(* IEC 61131-3 sources: codesys_asrs/Project_ASRS_CodeSYS (part 2) *)

(* ---- 16_FB_G3_Cycle_BODY_ONLY.st ---- *)
T_Nettoyage15(IN := NettoyageTimerEnable AND NOT GVL_SIG.ZONE_CONFIRMEE, PT := T#15m);
T_Prolong5(IN := ProlongTimerEnable AND NOT GVL_SIG.ZONE_CONFIRMEE, PT := T#5m);

// â”€â”€ Surveillance AU pendant cycle (prioritÃ© absolue) â”€â”€â”€â”€â”€â”€â”€â”€â”€â”€
IF GVL_SIG.OP_AU AND Step > 0 AND Step < 200 THEN
    GVL_SIG.G3_DEFAUT      := TRUE;
    GVL_SIG.G3_CODE_DEFAUT := 14;
    GVL_SEQ.DEFAUT_ACTIF   := TRUE;
    GVL_SEQ.CODE_DEFAUT    := 14;
    GVL_SIG.G4_REQ         := FALSE;
    GVL_SIG.G5_REQ         := FALSE;
    GVL_SIG.G6_REQ         := FALSE;
    GVL_SIG.G7_REQ         := FALSE;
    GVL_SIG.G8_REQ         := FALSE;
    GVL_SIG.G9_REQ_ARRET     := FALSE;
    GVL_SIG.G10_REQ_ENTRER   := FALSE;
    GVL_SIG.G10_REQ_SORTIR   := FALSE;
    GVL_SIG.VYT_CYCLE_EN_COURS := FALSE;
    Step := 0;
    RETURN;
END_IF;

CASE Step OF

// â•â•â•â•â•â•â•â•â•â•â•â•â•â•â•â•â•â•â•â•â•â•â•â•â•â•â•â•â•â•â•â•â•â•â•â•â•â•â•â•â•â•â•â•â•â•â•â•â•â•â•â•â•â•â•â•â•â•â•â•
// PHASE 0 â€” IDLE
// â•â•â•â•â•â•â•â•â•â•â•â•â•â•â•â•â•â•â•â•â•â•â•â•â•â•â•â•â•â•â•â•â•â•â•â•â•â•â•â•â•â•â•â•â•â•â•â•â•â•â•â•â•â•â•â•â•â•â•â•
0:
    GVL_SIG.G3_FIN_CM          := FALSE;
    GVL_SIG.G3_DEFAUT          := FALSE;
    GVL_SIG.G3_CODE_DEFAUT     := 0;
    GVL_SIG.VYT_CYCLE_EN_COURS := FALSE;
    GVL_SIG.G9_ARRETEE_OK      := FALSE;
    GVL_SIG.G9_DEBRIDE_OK      := FALSE;
    GVL_SIG.G9_BRIDE_OK        := FALSE;
    GVL_SIG.G9_AUTORISE_OK     := FALSE;
    GVL_SIG.G10_EN_PRESSE      := FALSE;
    GVL_SIG.G10_A_ZPM          := FALSE;
    NettoyageTimerEnable       := FALSE;
    ProlongTimerEnable         := FALSE;
    GVL_SIG.NETTOYAGE_EN_COURS := FALSE;
    GVL_SIG.NETTOYAGE_TIMEOUT  := FALSE;
    GVL_SIG.NETTOYAGE_PROLONGATION_UTILISEE := FALSE;
    GVL_SIG.NETTOYAGE_DEPASSEMENT_MAX := FALSE;
    GVL_SIG.VYT_NETTOYAGE_TIMEOUT := FALSE;
    GVL_IO.VOYANT_NETTOYAGE_TIMEOUT := FALSE;
    GVL_IO.VOYANT_NETTOYAGE_MAX := FALSE;
    GVL_IO.BUZZER_ATTENTE_ZONE_LIBRE := FALSE;
    IF GVL_SIG.G3_REQ THEN
        DepotFound := FALSE;
        PriseFound := FALSE;
        IF GVL_MOULES.MOULE_EN_PRESSE = 0 THEN
            GVL_SIG.G3_CODE_DEFAUT := 16;
            Step := 200;
        ELSIF GVL_MOULES.MOULE_DEMANDE = 0 THEN
            GVL_SIG.G3_CODE_DEFAUT := 13;
            Step := 200;
        ELSIF GVL_MOULES.MOULE_DEMANDE = GVL_MOULES.MOULE_EN_PRESSE THEN
            GVL_SIG.G3_CODE_DEFAUT := 17;
            Step := 200;
        ELSE
            Step := 1;
        END_IF;
    END_IF;

1: // Recherche slot dÃ©pÃ´t
    DepotFound := FALSE;
    FOR i := 1 TO 5 BY 1 DO
        IF NOT DepotFound THEN
            FOR j := 1 TO 2 BY 1 DO
                IF NOT DepotFound
                   AND NOT GVL_MOULES.CH[i, j].OCCUPE
                   AND NOT GVL_MOULES.CH[i, j].RESERVE THEN
                    GVL_MOULES.CIBLE_DEPOT_CH := INT_TO_USINT(i);
                    GVL_MOULES.CIBLE_DEPOT_NV := INT_TO_USINT(j);
                    GVL_MOULES.CH[i, j].RESERVE := TRUE;
                    DepotFound := TRUE;
                END_IF;
            END_FOR;
        END_IF;
    END_FOR;
    IF DepotFound THEN
        Step := 2;
    ELSE
        GVL_MOULES.ALM_STOCK_PLEIN := TRUE;
        GVL_SIG.ALM_STOCK_PLEIN   := TRUE;
        GVL_SIG.G3_CODE_DEFAUT    := 12;
        Step := 200;
    END_IF;

2: // Recherche slot prise
    PriseFound := FALSE;
    FOR i := 1 TO 5 BY 1 DO
        IF NOT PriseFound THEN
            FOR j := 1 TO 2 BY 1 DO
                IF NOT PriseFound
                   AND GVL_MOULES.CH[i, j].OCCUPE
                   AND GVL_MOULES.CH[i, j].ID = GVL_MOULES.MOULE_DEMANDE THEN
                    GVL_MOULES.CIBLE_PRISE_CH := INT_TO_USINT(i);
                    GVL_MOULES.CIBLE_PRISE_NV := INT_TO_USINT(j);
                    PriseFound := TRUE;
                END_IF;
            END_FOR;
        END_IF;
    END_FOR;
    IF PriseFound THEN
        GVL_SIG.VYT_CYCLE_EN_COURS := TRUE;
        Step := 3;
    ELSE
        GVL_MOULES.CH[GVL_MOULES.CIBLE_DEPOT_CH, GVL_MOULES.CIBLE_DEPOT_NV].RESERVE := FALSE;
        GVL_SIG.G3_CODE_DEFAUT := 13;
        Step := 200;
    END_IF;

3:
    GVL_SEQ.CYCLE_INTERROMPU := TRUE;
    GVL_SEQ.CYCLE_EN_COURS   := TRUE;

// â•â•â•â•â•â•â•â•â•â•â•â•â•â•â•â•â•â•â•â•â•â•â•â•â•â•â•â•â•â•â•â•â•â•â•â•â•â•â•â•â•â•â•â•â•â•â•â•â•â•â•â•â•â•â•â•â•â•â•â•
// PHASE 1 â€” ArrÃªt presse + dÃ©bridage
// â•â•â•â•â•â•â•â•â•â•â•â•â•â•â•â•â•â•â•â•â•â•â•â•â•â•â•â•â•â•â•â•â•â•â•â•â•â•â•â•â•â•â•â•â•â•â•â•â•â•â•â•â•â•â•â•â•â•â•â•
10:
    GVL_SIG.G9_REQ_ARRET   := TRUE;
    GVL_SIG.G10_REQ_ENTRER := TRUE;
    Step := 11;

11:
    IF GVL_SIG.G9_ARRETEE_OK THEN
        GVL_SIG.G9_REQ_DEBRIDAGE := TRUE;
        Step := 12;
    ELSIF GVL_SIG.G9_DEFAUT THEN
        Step := 200;
    END_IF;

12:
    IF GVL_SIG.G9_DEBRIDE_OK THEN
        Step := 13;
    ELSIF GVL_SIG.G9_DEFAUT THEN
        Step := 200;
    END_IF;

// â•â•â•â•â•â•â•â•â•â•â•â•â•â•â•â•â•â•â•â•â•â•â•â•â•â•â•â•â•â•â•â•â•â•â•â•â•â•â•â•â•â•â•â•â•â•â•â•â•â•â•â•â•â•â•â•â•â•â•â•
// DIVERGENCE ET#1 â€” Retrait introducteur â€– Chariot â†’ P0
// â•â•â•â•â•â•â•â•â•â•â•â•â•â•â•â•â•â•â•â•â•â•â•â•â•â•â•â•â•â•â•â•â•â•â•â•â•â•â•â•â•â•â•â•â•â•â•â•â•â•â•â•â•â•â•â•â•â•â•â•
13:
    BrA_Done := FALSE;
    BrB_Done := FALSE;
    SubA     := 0;
    SubB     := 0;
    Step     := 14;

14:
    IF NOT BrA_Done THEN
        CASE SubA OF
        0:  GVL_SIG.G10_REQ_SORTIR := TRUE;
            SubA := 1;
        1:  IF GVL_SIG.G10_A_ZPM THEN
                BrA_Done := TRUE;
            ELSIF GVL_SIG.G10_DEFAUT THEN
                GVL_SIG.G3_CODE_DEFAUT := 5;
                Step := 200;
            END_IF;
        END_CASE;
    END_IF;

    IF NOT BrB_Done THEN
        CASE SubB OF
        0:  GVL_SIG.G4_REQ   := TRUE;
            GVL_SIG.G4_CIBLE := 0;
            SubB := 1;
        1:  IF GVL_SIG.G4_DONE THEN
                GVL_SIG.G4_DONE := FALSE;
                BrB_Done := TRUE;
            ELSIF GVL_SIG.G4_ERR THEN
                GVL_SIG.G4_ERR := FALSE;
                GVL_SIG.G3_CODE_DEFAUT := 7;
                Step := 200;
            END_IF;
        END_CASE;
    END_IF;

    IF BrA_Done AND BrB_Done THEN
        GVL_SIG.G10_REQ_ENTRER := FALSE;
        GVL_SIG.G10_REQ_SORTIR := FALSE;
        Step := 15;
    END_IF;

// â•â•â•â•â•â•â•â•â•â•â•â•â•â•â•â•â•â•â•â•â•â•â•â•â•â•â•â•â•â•â•â•â•â•â•â•â•â•â•â•â•â•â•â•â•â•â•â•â•â•â•â•â•â•â•â•â•â•â•â•
// PHASE 2 â€” Transfert moule : introducteur â†’ chariot
// â•â•â•â•â•â•â•â•â•â•â•â•â•â•â•â•â•â•â•â•â•â•â•â•â•â•â•â•â•â•â•â•â•â•â•â•â•â•â•â•â•â•â•â•â•â•â•â•â•â•â•â•â•â•â•â•â•â•â•â•
15:
    IF NOT GVL_IO.MOULE_SUR_INTRO THEN
        GVL_SIG.G3_CODE_DEFAUT := 13;
        Step := 200;
    ELSE
        Step := 16;
    END_IF;

16:
    GVL_SIG.G6_REQ   := TRUE;
    GVL_SIG.G6_CIBLE := 0;  // NORD
    Step := 17;

17:
    IF GVL_SIG.G6_DONE THEN
        GVL_SIG.G6_DONE := FALSE;
        Step := 18;
    ELSIF GVL_SIG.G6_ERR THEN
        GVL_SIG.G6_ERR         := FALSE;
        GVL_SIG.G3_CODE_DEFAUT := 11;
        Step := 200;
    END_IF;

18:
    GVL_SIG.G5_REQ   := TRUE;
    GVL_SIG.G5_CIBLE := 0;  // Z_ZPM
    Step := 19;

19:
    IF GVL_SIG.G5_DONE THEN
        GVL_SIG.G5_DONE := FALSE;
        Step := 20;
    ELSIF GVL_SIG.G5_ERR THEN
        GVL_SIG.G5_ERR         := FALSE;
        GVL_SIG.G3_CODE_DEFAUT := 6;
        Step := 200;
    END_IF;

20:
    GVL_SIG.G7_REQ := TRUE;
    GVL_SIG.G7_CMD := 0;  // ETENDRE
    Step := 21;

21:
    IF GVL_SIG.G7_DONE THEN
        GVL_SIG.G7_DONE := FALSE;
        Step := 22;
    ELSIF GVL_SIG.G7_ERR THEN
        GVL_SIG.G7_ERR         := FALSE;
        GVL_SIG.G3_CODE_DEFAUT := 11;
        Step := 200;
    END_IF;

22:
    GVL_SIG.G5_REQ   := TRUE;
    GVL_SIG.G5_CIBLE := 3;  // Z_TRANSPORT
    Step := 23;

23:
    IF GVL_SIG.G5_DONE THEN
        GVL_SIG.G5_DONE := FALSE;
        IF NOT GVL_IO.CAPTEUR_CHARGE_CHARIOT THEN
            GVL_SIG.G3_CODE_DEFAUT := 10;
            Step := 200;
        ELSE
            Step := 24;
        END_IF;
    ELSIF GVL_SIG.G5_ERR THEN
        GVL_SIG.G5_ERR         := FALSE;
        GVL_SIG.G3_CODE_DEFAUT := 6;
        Step := 200;
    END_IF;

24:
    GVL_SIG.G7_REQ := TRUE;
    GVL_SIG.G7_CMD := 1;  // RETRACTER
    Step := 25;

25:
    IF GVL_SIG.G7_DONE THEN
        GVL_SIG.G7_DONE := FALSE;
        Step := 26;
    ELSIF GVL_SIG.G7_ERR THEN
        GVL_SIG.G7_ERR         := FALSE;
        GVL_SIG.G3_CODE_DEFAUT := 11;
        Step := 201;
    END_IF;

// â•â•â•â•â•â•â•â•â•â•â•â•â•â•â•â•â•â•â•â•â•â•â•â•â•â•â•â•â•â•â•â•â•â•â•â•â•â•â•â•â•â•â•â•â•â•â•â•â•â•â•â•â•â•â•â•â•â•â•â•
// DIVERGENCE ET#2 â€” Stockage+RFID+Prise â€– Nettoyage
// â•â•â•â•â•â•â•â•â•â•â•â•â•â•â•â•â•â•â•â•â•â•â•â•â•â•â•â•â•â•â•â•â•â•â•â•â•â•â•â•â•â•â•â•â•â•â•â•â•â•â•â•â•â•â•â•â•â•â•â•
26:
    BrA_Done := FALSE;
    BrB_Done := FALSE;
    SubA     := 0;
    SubB     := 0;
    NettoyageTimerEnable := FALSE;
    ProlongTimerEnable := FALSE;
    GVL_SIG.NETTOYAGE_EN_COURS := FALSE;
    GVL_SIG.NETTOYAGE_TIMEOUT := FALSE;
    GVL_SIG.NETTOYAGE_PROLONGATION_UTILISEE := FALSE;
    GVL_SIG.NETTOYAGE_DEPASSEMENT_MAX := FALSE;
    GVL_SIG.VYT_NETTOYAGE_TIMEOUT := FALSE;
    GVL_IO.VOYANT_NETTOYAGE_TIMEOUT := FALSE;
    GVL_IO.VOYANT_NETTOYAGE_MAX := FALSE;
    GVL_IO.BUZZER_ATTENTE_ZONE_LIBRE := FALSE;
    Step     := 27;

27: // ET#2
    IF NOT BrA_Done THEN
        CASE SubA OF
        0:  GVL_SIG.G4_REQ   := TRUE;
            GVL_SIG.G4_CIBLE := GVL_MOULES.CIBLE_DEPOT_CH;
            SubA := 1;
        1:  IF GVL_SIG.G4_DONE THEN
                GVL_SIG.G4_DONE := FALSE; SubA := 2;
            ELSIF GVL_SIG.G4_ERR THEN
                GVL_SIG.G4_ERR := FALSE;
                GVL_SIG.G3_CODE_DEFAUT := 7; Step := 201; END_IF;
        2:  GVL_SIG.G6_REQ   := TRUE;
            GVL_SIG.G6_CIBLE := 1; // SUD
            SubA := 3;
        3:  IF GVL_SIG.G6_DONE THEN
                GVL_SIG.G6_DONE := FALSE; SubA := 4;
            ELSIF GVL_SIG.G6_ERR THEN
                GVL_SIG.G6_ERR := FALSE;
                GVL_SIG.G3_CODE_DEFAUT := 11; Step := 201; END_IF;
        4:  GVL_SIG.G7_REQ := TRUE;
            GVL_SIG.G7_CMD := 0; // EXT
            SubA := 5;
        5:  IF GVL_SIG.G7_DONE THEN
                GVL_SIG.G7_DONE := FALSE; SubA := 6;
            ELSIF GVL_SIG.G7_ERR THEN
                GVL_SIG.G7_ERR := FALSE;
                GVL_SIG.G3_CODE_DEFAUT := 11; Step := 201; END_IF;
        6:  GVL_SIG.G5_REQ   := TRUE;
            GVL_SIG.G5_CIBLE := GVL_MOULES.CIBLE_DEPOT_NV;
            SubA := 7;
        7:  IF GVL_SIG.G5_DONE THEN
                GVL_SIG.G5_DONE := FALSE; SubA := 8;
            ELSIF GVL_SIG.G5_ERR THEN
                GVL_SIG.G5_ERR := FALSE;
                GVL_SIG.G3_CODE_DEFAUT := 6; Step := 201; END_IF;
        8:  GVL_SIG.G7_REQ := TRUE;
            GVL_SIG.G7_CMD := 1; // RET
            SubA := 9;
        9:  IF GVL_SIG.G7_DONE THEN
                GVL_SIG.G7_DONE := FALSE;
                IF NOT GVL_SIG.CAPTEUR_PRES_CH[GVL_MOULES.CIBLE_DEPOT_CH,
                                               GVL_MOULES.CIBLE_DEPOT_NV] THEN
                    GVL_SIG.G3_CODE_DEFAUT := 11; Step := 202;
                ELSE
                    GVL_MOULES.CH[GVL_MOULES.CIBLE_DEPOT_CH,
                                  GVL_MOULES.CIBLE_DEPOT_NV].OCCUPE  := TRUE;
                    GVL_MOULES.CH[GVL_MOULES.CIBLE_DEPOT_CH,
                                  GVL_MOULES.CIBLE_DEPOT_NV].ID      := GVL_MOULES.MOULE_EN_PRESSE;
                    GVL_MOULES.CH[GVL_MOULES.CIBLE_DEPOT_CH,
                                  GVL_MOULES.CIBLE_DEPOT_NV].RESERVE := FALSE;
                    IF GVL_MOULES.NB_EMPLACEMENTS_LIBRES > 0 THEN
                        GVL_MOULES.NB_EMPLACEMENTS_LIBRES :=
                            GVL_MOULES.NB_EMPLACEMENTS_LIBRES - 1;
                    END_IF;
                    SubA := 10;
                END_IF;
            ELSIF GVL_SIG.G7_ERR THEN
                GVL_SIG.G7_ERR := FALSE;
                GVL_SIG.G3_CODE_DEFAUT := 11; Step := 202; END_IF;
        10: GVL_SIG.G5_REQ   := TRUE;
            GVL_SIG.G5_CIBLE := 3; // Z_TRANSPORT
            SubA := 11;
        11: IF GVL_SIG.G5_DONE THEN
                GVL_SIG.G5_DONE := FALSE; SubA := 12;
            ELSIF GVL_SIG.G5_ERR THEN
                GVL_SIG.G5_ERR := FALSE;
                GVL_SIG.G3_CODE_DEFAUT := 6; Step := 202; END_IF;
        12: GVL_SIG.G4_REQ   := TRUE;
            GVL_SIG.G4_CIBLE := GVL_MOULES.CIBLE_PRISE_CH;
            SubA := 13;
        13: IF GVL_SIG.G4_DONE THEN
                GVL_SIG.G4_DONE := FALSE; SubA := 14;
            ELSIF GVL_SIG.G4_ERR THEN
                GVL_SIG.G4_ERR := FALSE;
                GVL_SIG.G3_CODE_DEFAUT := 7; Step := 202; END_IF;
        14: GVL_SIG.G8_REQ        := TRUE;
            GVL_SIG.G8_ID_ATTENDU := GVL_MOULES.MOULE_DEMANDE;
            SubA := 15;
        15: IF GVL_SIG.G8_DONE THEN
                GVL_SIG.G8_DONE := FALSE;
                IF GVL_SIG.G8_OK THEN
                    GVL_MOULES.CH[GVL_MOULES.CIBLE_PRISE_CH,
                                  GVL_MOULES.CIBLE_PRISE_NV].RFID_OK := TRUE;
                    SubA := 16;
                ELSE
                    GVL_SIG.G8_ERR         := FALSE;
                    GVL_SIG.G3_CODE_DEFAUT := 8;
                    Step := 202;
                END_IF;
            ELSIF GVL_SIG.G8_ERR THEN
                GVL_SIG.G8_ERR         := FALSE;
                GVL_SIG.G3_CODE_DEFAUT := 8; Step := 202; END_IF;
        16: GVL_SIG.G5_REQ   := TRUE;
            GVL_SIG.G5_CIBLE := GVL_MOULES.CIBLE_PRISE_NV;
            SubA := 17;
        17: IF GVL_SIG.G5_DONE THEN
                GVL_SIG.G5_DONE := FALSE; SubA := 18;
            ELSIF GVL_SIG.G5_ERR THEN
                GVL_SIG.G5_ERR := FALSE;
                GVL_SIG.G3_CODE_DEFAUT := 6; Step := 202; END_IF;
        18: GVL_SIG.G7_REQ := TRUE;
            GVL_SIG.G7_CMD := 0; // EXT
            SubA := 19;
        19: IF GVL_SIG.G7_DONE THEN
                GVL_SIG.G7_DONE := FALSE; SubA := 20;
            ELSIF GVL_SIG.G7_ERR THEN
                GVL_SIG.G7_ERR := FALSE;
                GVL_SIG.G3_CODE_DEFAUT := 11; Step := 202; END_IF;
        20: GVL_SIG.G5_REQ   := TRUE;
            GVL_SIG.G5_CIBLE := 3; // Z_TRANSPORT
            SubA := 21;
        21: IF GVL_SIG.G5_DONE THEN
                GVL_SIG.G5_DONE := FALSE;
                IF NOT GVL_IO.CAPTEUR_CHARGE_CHARIOT THEN
                    GVL_SIG.G3_CODE_DEFAUT := 10; Step := 202;
                ELSE
                    SubA := 22;
                END_IF;
            ELSIF GVL_SIG.G5_ERR THEN
                GVL_SIG.G5_ERR := FALSE;
                GVL_SIG.G3_CODE_DEFAUT := 6; Step := 202; END_IF;
        22: GVL_SIG.G7_REQ := TRUE;
            GVL_SIG.G7_CMD := 1; // RET
            SubA := 23;
        23: IF GVL_SIG.G7_DONE THEN
                GVL_SIG.G7_DONE := FALSE;
                GVL_MOULES.CH[GVL_MOULES.CIBLE_PRISE_CH,
                               GVL_MOULES.CIBLE_PRISE_NV].OCCUPE := FALSE;
                GVL_MOULES.CH[GVL_MOULES.CIBLE_PRISE_CH,
                               GVL_MOULES.CIBLE_PRISE_NV].ID     := 0;
                GVL_MOULES.NB_EMPLACEMENTS_LIBRES :=
                    GVL_MOULES.NB_EMPLACEMENTS_LIBRES + 1;
                GVL_SEQ.MOULE_EN_TRANSIT := TRUE;
                SubA := 24;
            ELSIF GVL_SIG.G7_ERR THEN
                GVL_SIG.G7_ERR := FALSE;
                GVL_SIG.G3_CODE_DEFAUT := 11; Step := 203; END_IF;
        24: GVL_SIG.G4_REQ   := TRUE;
            GVL_SIG.G4_CIBLE := 0; // P0
            SubA := 25;
        25: IF GVL_SIG.G4_DONE THEN
                GVL_SIG.G4_DONE := FALSE; SubA := 26;
            ELSIF GVL_SIG.G4_ERR THEN
                GVL_SIG.G4_ERR := FALSE;
                GVL_SIG.G3_CODE_DEFAUT := 7; Step := 203; END_IF;
        26: GVL_SIG.G8_REQ        := TRUE;
            GVL_SIG.G8_ID_ATTENDU := GVL_MOULES.MOULE_DEMANDE;
            SubA := 27;
        27: IF GVL_SIG.G8_DONE THEN
                GVL_SIG.G8_DONE := FALSE;
                IF GVL_SIG.G8_OK THEN
                    BrA_Done := TRUE;
                ELSE
                    GVL_SIG.G8_ERR         := FALSE;
                    GVL_SIG.G3_CODE_DEFAUT := 9;
                    Step := 210;
                END_IF;
            ELSIF GVL_SIG.G8_ERR THEN
                GVL_SIG.G8_ERR         := FALSE;
                GVL_SIG.G3_CODE_DEFAUT := 9; Step := 210; END_IF;
        END_CASE;
    END_IF;

    IF NOT BrB_Done THEN
        CASE SubB OF
        0:  GVL_SIG.VYT_NETTOYAGE  := TRUE;
            GVL_IO.VOYANT_NETTOYAGE := TRUE;
            IF SubA >= 10 THEN
                GVL_IO.BUZZER_DEBUT_NETTOYAGE := TRUE;
                NettoyageTimerEnable := TRUE;
                ProlongTimerEnable := FALSE;
                GVL_SIG.NETTOYAGE_EN_COURS := TRUE;
                GVL_SIG.NETTOYAGE_TIMEOUT := FALSE;
                GVL_SIG.NETTOYAGE_PROLONGATION_UTILISEE := FALSE;
                GVL_SIG.NETTOYAGE_DEPASSEMENT_MAX := FALSE;
                SubB := 1;
            END_IF;

        1:  GVL_IO.BUZZER_DEBUT_NETTOYAGE := FALSE;
            GVL_SIG.VYT_ATTENTE_ZONE := NOT GVL_SIG.ZONE_CONFIRMEE;
            GVL_IO.VOYANT_ATTENTE_ZONE_LIBRE := NOT GVL_SIG.ZONE_CONFIRMEE;

            IF GVL_SIG.ZONE_CONFIRMEE THEN
                GVL_IO.VOYANT_NETTOYAGE := FALSE;
                GVL_IO.VOYANT_ATTENTE_ZONE_LIBRE := FALSE;
                GVL_IO.VOYANT_NETTOYAGE_TIMEOUT := FALSE;
                GVL_IO.VOYANT_NETTOYAGE_MAX := FALSE;
                GVL_IO.BUZZER_ATTENTE_ZONE_LIBRE := FALSE;
                GVL_SIG.VYT_NETTOYAGE := FALSE;
                GVL_SIG.VYT_ATTENTE_ZONE := FALSE;
                GVL_SIG.VYT_NETTOYAGE_TIMEOUT := FALSE;
                GVL_SIG.NETTOYAGE_EN_COURS := FALSE;
                GVL_SIG.NETTOYAGE_TIMEOUT := FALSE;
                NettoyageTimerEnable := FALSE;
                ProlongTimerEnable := FALSE;
                BrB_Done := TRUE;

            ELSIF T_Prolong5.Q THEN
                GVL_SIG.NETTOYAGE_DEPASSEMENT_MAX := TRUE;
                GVL_SIG.NETTOYAGE_TIMEOUT := TRUE;
                GVL_SIG.VYT_NETTOYAGE_TIMEOUT := TRUE;
                GVL_IO.VOYANT_NETTOYAGE_TIMEOUT := TRUE;
                GVL_IO.VOYANT_NETTOYAGE_MAX := TRUE;
                GVL_IO.BUZZER_ATTENTE_ZONE_LIBRE := TRUE;
                GVL_SIG.G3_CODE_DEFAUT := 18;
                IF GVL_SEQ.MOULE_EN_TRANSIT THEN
                    Step := 203;
                ELSE
                    Step := 202;
                END_IF;

            ELSIF T_Nettoyage15.Q THEN
                GVL_SIG.NETTOYAGE_TIMEOUT := TRUE;
                GVL_SIG.VYT_NETTOYAGE_TIMEOUT := TRUE;
                GVL_IO.VOYANT_NETTOYAGE_TIMEOUT := TRUE;
                GVL_IO.BUZZER_ATTENTE_ZONE_LIBRE := TRUE;

                IF GVL_SIG.OP_PROLONG_NETTOYAGE
                   AND NOT GVL_SIG.NETTOYAGE_PROLONGATION_UTILISEE THEN
                    GVL_SIG.NETTOYAGE_PROLONGATION_UTILISEE := TRUE;
                    GVL_SIG.NETTOYAGE_TIMEOUT := FALSE;
                    GVL_SIG.VYT_NETTOYAGE_TIMEOUT := FALSE;
                    GVL_IO.VOYANT_NETTOYAGE_TIMEOUT := FALSE;
                    GVL_IO.BUZZER_ATTENTE_ZONE_LIBRE := FALSE;
                    NettoyageTimerEnable := FALSE;
                    ProlongTimerEnable := TRUE;
                END_IF;
            END_IF;
        END_CASE;
    END_IF;

    IF BrA_Done AND BrB_Done THEN
        Step := 30;
    END_IF;

// â•â•â•â•â•â•â•â•â•â•â•â•â•â•â•â•â•â•â•â•â•â•â•â•â•â•â•â•â•â•â•â•â•â•â•â•â•â•â•â•â•â•â•â•â•â•â•â•â•â•â•â•â•â•â•â•â•â•â•â•
// PHASE 3 â€” DÃ©pÃ´t nouveau moule sur introducteur
// â•â•â•â•â•â•â•â•â•â•â•â•â•â•â•â•â•â•â•â•â•â•â•â•â•â•â•â•â•â•â•â•â•â•â•â•â•â•â•â•â•â•â•â•â•â•â•â•â•â•â•â•â•â•â•â•â•â•â•â•
30:
    GVL_SIG.G6_REQ   := TRUE;
    GVL_SIG.G6_CIBLE := 0; // NORD
    Step := 31;

31:
    IF GVL_SIG.G6_DONE THEN
        GVL_SIG.G6_DONE := FALSE; Step := 32;
    ELSIF GVL_SIG.G6_ERR THEN
        GVL_SIG.G6_ERR         := FALSE;
        GVL_SIG.G3_CODE_DEFAUT := 11; Step := 203; END_IF;

32:
    GVL_SIG.G7_REQ := TRUE;
    GVL_SIG.G7_CMD := 0; // EXT
    Step := 33;

33:
    IF GVL_SIG.G7_DONE THEN
        GVL_SIG.G7_DONE := FALSE; Step := 34;
    ELSIF GVL_SIG.G7_ERR THEN
        GVL_SIG.G7_ERR         := FALSE;
        GVL_SIG.G3_CODE_DEFAUT := 11; Step := 203; END_IF;

34:
    GVL_SIG.G5_REQ   := TRUE;
    GVL_SIG.G5_CIBLE := 0; // Z_ZPM
    Step := 35;

35:
    IF GVL_SIG.G5_DONE THEN
        GVL_SIG.G5_DONE := FALSE; Step := 36;
    ELSIF GVL_SIG.G5_ERR THEN
        GVL_SIG.G5_ERR         := FALSE;
        GVL_SIG.G3_CODE_DEFAUT := 6; Step := 203; END_IF;

36:
    GVL_SIG.G7_REQ := TRUE;
    GVL_SIG.G7_CMD := 1; // RET
    Step := 37;

37:
    IF GVL_SIG.G7_DONE THEN
        GVL_SIG.G7_DONE := FALSE;
        IF NOT GVL_IO.MOULE_SUR_INTRO THEN
            GVL_SIG.G3_CODE_DEFAUT := 11; Step := 203;
        ELSIF GVL_IO.CAPTEUR_CHARGE_CHARIOT THEN
            GVL_SIG.G3_CODE_DEFAUT := 11; Step := 203;
        ELSE
            Step := 38;
        END_IF;
    ELSIF GVL_SIG.G7_ERR THEN
        GVL_SIG.G7_ERR         := FALSE;
        GVL_SIG.G3_CODE_DEFAUT := 11; Step := 203; END_IF;

38:
    GVL_SIG.G5_REQ   := TRUE;
    GVL_SIG.G5_CIBLE := 3; // Z_TRANSPORT
    Step := 39;

39:
    IF GVL_SIG.G5_DONE THEN
        GVL_SIG.G5_DONE         := FALSE;
        GVL_SIG.G10_REQ_ENTRER  := TRUE;
        GVL_SIG.G9_REQ_BRIDAGE  := TRUE;
        Step := 40;
    ELSIF GVL_SIG.G5_ERR THEN
        GVL_SIG.G5_ERR         := FALSE;
        GVL_SIG.G3_CODE_DEFAUT := 6; Step := 203; END_IF;

40:
    IF GVL_SIG.G9_BRIDE_OK AND GVL_SIG.G10_A_ZPM THEN
        GVL_MOULES.MOULE_EN_PRESSE := GVL_MOULES.MOULE_DEMANDE;
        GVL_SEQ.MOULE_EN_TRANSIT   := FALSE;
        GVL_SIG.G10_REQ_ENTRER     := FALSE;
        Step := 41;
    ELSIF GVL_SIG.G9_DEFAUT THEN
        GVL_SIG.G3_CODE_DEFAUT := 3; Step := 200;
    ELSIF GVL_SIG.G10_DEFAUT THEN
        GVL_SIG.G3_CODE_DEFAUT := 5; Step := 200;
    END_IF;

// â•â•â•â•â•â•â•â•â•â•â•â•â•â•â•â•â•â•â•â•â•â•â•â•â•â•â•â•â•â•â•â•â•â•â•â•â•â•â•â•â•â•â•â•â•â•â•â•â•â•â•â•â•â•â•â•â•â•â•â•
// DIVERGENCE ET#3 â€” Autorisation presse â€– Retour garage
// â•â•â•â•â•â•â•â•â•â•â•â•â•â•â•â•â•â•â•â•â•â•â•â•â•â•â•â•â•â•â•â•â•â•â•â•â•â•â•â•â•â•â•â•â•â•â•â•â•â•â•â•â•â•â•â•â•â•â•â•
41:
    BrA_Done := FALSE;
    BrB_Done := FALSE;
    SubA     := 0;
    SubB     := 0;
    Step     := 42;

42:
    IF NOT BrA_Done THEN
        CASE SubA OF
        0:  GVL_SIG.G9_REQ_AUTORISER := TRUE;
            SubA := 1;
        1:  IF GVL_SIG.G9_AUTORISE_OK THEN
                GVL_SIG.G9_REQ_AUTORISER := FALSE;
                BrA_Done := TRUE;
            ELSIF GVL_SIG.G9_DEFAUT THEN
                GVL_SIG.G3_CODE_DEFAUT := 3; Step := 200; END_IF;
        END_CASE;
    END_IF;

    IF NOT BrB_Done THEN
        CASE SubB OF
        0:  GVL_SIG.G4_REQ   := TRUE;
            GVL_SIG.G4_CIBLE := 6; // P6 Garage
            SubB := 1;
        1:  IF GVL_SIG.G4_DONE THEN
                GVL_SIG.G4_DONE := FALSE;
                BrB_Done := TRUE;
            ELSIF GVL_SIG.G4_ERR THEN
                GVL_SIG.G4_ERR := FALSE;
                BrB_Done := TRUE;  // Non bloquant
            END_IF;
        END_CASE;
    END_IF;

    IF BrA_Done AND BrB_Done THEN
        Step := 50;
    END_IF;

// â•â•â•â•â•â•â•â•â•â•â•â•â•â•â•â•â•â•â•â•â•â•â•â•â•â•â•â•â•â•â•â•â•â•â•â•â•â•â•â•â•â•â•â•â•â•â•â•â•â•â•â•â•â•â•â•â•â•â•â•
// PHASE FINALE â€” Fin de cycle
// â•â•â•â•â•â•â•â•â•â•â•â•â•â•â•â•â•â•â•â•â•â•â•â•â•â•â•â•â•â•â•â•â•â•â•â•â•â•â•â•â•â•â•â•â•â•â•â•â•â•â•â•â•â•â•â•â•â•â•â•
50:
    GVL_SEQ.CYCLE_INTERROMPU    := FALSE;
    GVL_SEQ.CYCLE_EN_COURS      := FALSE;
    GVL_MOULES.ALM_STOCK_PLEIN  := FALSE;
    GVL_SIG.VYT_CYCLE_EN_COURS  := FALSE;
    GVL_SIG.G3_FIN_CM           := TRUE;
    IF NOT GVL_SIG.G3_REQ THEN
        GVL_SIG.G3_FIN_CM := FALSE;
        Step := 0;
    END_IF;

// â•â•â•â•â•â•â•â•â•â•â•â•â•â•â•â•â•â•â•â•â•â•â•â•â•â•â•â•â•â•â•â•â•â•â•â•â•â•â•â•â•â•â•â•â•â•â•â•â•â•â•â•â•â•â•â•â•â•â•â•
// BRANCHES DÃ‰FAUT
// â•â•â•â•â•â•â•â•â•â•â•â•â•â•â•â•â•â•â•â•â•â•â•â•â•â•â•â•â•â•â•â•â•â•â•â•â•â•â•â•â•â•â•â•â•â•â•â•â•â•â•â•â•â•â•â•â•â•â•â•
200: // DÃ©faut chariot VIDE
    GVL_SIG.G3_DEFAUT          := TRUE;
    GVL_SEQ.DEFAUT_ACTIF       := TRUE;
    GVL_SEQ.CODE_DEFAUT        := GVL_SIG.G3_CODE_DEFAUT;
    GVL_SIG.VYT_CYCLE_EN_COURS := FALSE;
    GVL_SIG.VYT_DEFAUT         := TRUE;
    IF GVL_MOULES.CIBLE_DEPOT_CH >= 1
       AND GVL_MOULES.CIBLE_DEPOT_CH <= 5 THEN
        GVL_MOULES.CH[GVL_MOULES.CIBLE_DEPOT_CH,
                      GVL_MOULES.CIBLE_DEPOT_NV].RESERVE := FALSE;
    END_IF;
    IF GVL_SIG.OP_CMD_RESET AND GVL_SIG.OP_CMD_ACQ THEN
        GVL_SIG.G3_DEFAUT    := FALSE;
        GVL_SEQ.DEFAUT_ACTIF := FALSE;
        GVL_SEQ.CODE_DEFAUT  := 0;
        GVL_SIG.VYT_DEFAUT   := FALSE;
        GVL_SEQ.CYCLE_INTERROMPU := FALSE;
        Step := 0;
    END_IF;

201: // DÃ©faut ancien moule sur fourches
    GVL_SIG.G3_DEFAUT          := TRUE;
    GVL_SEQ.DEFAUT_ACTIF       := TRUE;
    GVL_SEQ.CODE_DEFAUT        := GVL_SIG.G3_CODE_DEFAUT;
    GVL_SIG.VYT_DEFAUT         := TRUE;
    GVL_SIG.VYT_CYCLE_EN_COURS := FALSE;
    IF GVL_SIG.OP_CMD_RESET AND GVL_SIG.OP_CMD_ACQ THEN
        GVL_SIG.G3_DEFAUT    := FALSE;
        GVL_SEQ.DEFAUT_ACTIF := FALSE;
        GVL_SIG.VYT_DEFAUT   := FALSE;
        Step := 0;
    END_IF;

202: // DÃ©faut ancien moule dÃ©posÃ©, chariot vide
    GVL_SIG.G3_DEFAUT          := TRUE;
    GVL_SEQ.DEFAUT_ACTIF       := TRUE;
    GVL_SEQ.CODE_DEFAUT        := GVL_SIG.G3_CODE_DEFAUT;
    GVL_SIG.VYT_DEFAUT         := TRUE;
    GVL_SIG.VYT_CYCLE_EN_COURS := FALSE;
    IF GVL_SIG.OP_CMD_RESET AND GVL_SIG.OP_CMD_ACQ THEN
        GVL_SIG.G3_DEFAUT    := FALSE;
        GVL_SEQ.DEFAUT_ACTIF := FALSE;
        GVL_SIG.VYT_DEFAUT   := FALSE;
        Step := 0;
    END_IF;

203: // DÃ©faut nouveau moule sur fourches (MOULE_EN_TRANSIT=TRUE)
    GVL_SIG.G3_DEFAUT          := TRUE;
    GVL_SEQ.DEFAUT_ACTIF       := TRUE;
    GVL_SEQ.CODE_DEFAUT        := GVL_SIG.G3_CODE_DEFAUT;
    GVL_SIG.VYT_DEFAUT         := TRUE;
    GVL_SIG.VYT_CYCLE_EN_COURS := FALSE;
    IF GVL_SIG.OP_CMD_RESET AND GVL_SIG.OP_CMD_ACQ THEN
        GVL_SIG.G3_DEFAUT    := FALSE;
        GVL_SEQ.DEFAUT_ACTIF := FALSE;
        GVL_SIG.VYT_DEFAUT   := FALSE;
        Step := 0;
    END_IF;

210: // RFID2 KO â€” ROLLBACK (remettre moule en chambre prise)
    GVL_SIG.ALM_RFID           := TRUE;
    GVL_SIG.G3_DEFAUT          := TRUE;
    GVL_SEQ.DEFAUT_ACTIF       := TRUE;
    GVL_SEQ.CODE_DEFAUT        := 9;
    GVL_SIG.VYT_CYCLE_EN_COURS := FALSE;
    GVL_SIG.VYT_DEFAUT         := TRUE;
    GVL_MOULES.CH[GVL_MOULES.CIBLE_PRISE_CH,
                  GVL_MOULES.CIBLE_PRISE_NV].OCCUPE := TRUE;
    GVL_MOULES.CH[GVL_MOULES.CIBLE_PRISE_CH,
                  GVL_MOULES.CIBLE_PRISE_NV].ID     := GVL_MOULES.MOULE_DEMANDE;
    GVL_MOULES.NB_EMPLACEMENTS_LIBRES :=
        GVL_MOULES.NB_EMPLACEMENTS_LIBRES - 1;
    GVL_SEQ.MOULE_EN_TRANSIT := FALSE;
    IF GVL_SIG.OP_CMD_RESET AND GVL_SIG.OP_CMD_ACQ THEN
        GVL_SIG.G3_DEFAUT    := FALSE;
        GVL_SEQ.DEFAUT_ACTIF := FALSE;
        GVL_SIG.ALM_RFID     := FALSE;
        GVL_SIG.VYT_DEFAUT   := FALSE;
        Step := 0;
    END_IF;

END_CASE;

(* ---- 17_PRG_STARTUP.st ---- *)
// ================================================================
// 17_PRG_STARTUP.st  —  Programme démarrage (équivalent OB100)
// CODESYS V3.5 — PROGRAM
// Configurer cette tâche en "Single" dans le Task Manager CODESYS
// (exécution une seule fois au démarrage)
// ================================================================

PROGRAM PRG_STARTUP
VAR
END_VAR

// ── Initialisation GVL_SIG ────────────────────────────────────
GVL_SIG.SECURITES_OK        := FALSE;
GVL_SIG.ZONE_CONFIRMEE      := FALSE;
GVL_SIG.DEFAUT_AXE          := FALSE;
GVL_SIG.PERTE_PROFINET      := FALSE;
GVL_SIG.G2_REQ              := FALSE;
GVL_SIG.G2_HOMING_OK        := FALSE;
GVL_SIG.G2_DEFAUT           := FALSE;
GVL_SIG.G3_REQ              := FALSE;
GVL_SIG.G3_FIN_CM           := FALSE;
GVL_SIG.G3_DEFAUT           := FALSE;
GVL_SIG.G3_CODE_DEFAUT      := 0;
GVL_SIG.G4_REQ              := FALSE;
GVL_SIG.G4_DONE             := FALSE;
GVL_SIG.G4_ERR              := FALSE;
GVL_SIG.G5_REQ              := FALSE;
GVL_SIG.G5_DONE             := FALSE;
GVL_SIG.G5_ERR              := FALSE;
GVL_SIG.G6_REQ              := FALSE;
GVL_SIG.G6_DONE             := FALSE;
GVL_SIG.G6_ERR              := FALSE;
GVL_SIG.G7_REQ              := FALSE;
GVL_SIG.G7_DONE             := FALSE;
GVL_SIG.G7_ERR              := FALSE;
GVL_SIG.G8_REQ              := FALSE;
GVL_SIG.G8_DONE             := FALSE;
GVL_SIG.G8_OK               := FALSE;
GVL_SIG.G8_ERR              := FALSE;
GVL_SIG.G9_REQ_ARRET        := FALSE;
GVL_SIG.G9_REQ_DEBRIDAGE    := FALSE;
GVL_SIG.G9_REQ_BRIDAGE      := FALSE;
GVL_SIG.G9_REQ_AUTORISER    := FALSE;
GVL_SIG.G9_ARRETEE_OK       := FALSE;
GVL_SIG.G9_DEBRIDE_OK       := FALSE;
GVL_SIG.G9_BRIDE_OK         := FALSE;
GVL_SIG.G9_AUTORISE_OK      := FALSE;
GVL_SIG.G9_DEFAUT           := FALSE;
GVL_SIG.G10_REQ_ENTRER      := FALSE;
GVL_SIG.G10_REQ_SORTIR      := FALSE;
GVL_SIG.G10_EN_PRESSE       := FALSE;
GVL_SIG.G10_A_ZPM           := FALSE;
GVL_SIG.G10_DEFAUT          := FALSE;
GVL_SIG.VYT_MACHINE_PRETE   := FALSE;
GVL_SIG.VYT_CYCLE_EN_COURS  := FALSE;
GVL_SIG.VYT_DEFAUT          := FALSE;
GVL_SIG.VYT_INIT_OK         := FALSE;
GVL_SIG.CYCLE_CM_AUTORISE   := FALSE;

// ── Initialisation GVL_SEQ (hors Retain) ─────────────────────
// CYCLE_INTERROMPU, MOULE_EN_TRANSIT, NB_CYCLES_TOTAL = Retain → conservés
GVL_SEQ.ETAPE_ACTIVE    := 0;
GVL_SEQ.CYCLE_EN_COURS  := FALSE;
GVL_SEQ.HOMING_OK       := FALSE;
GVL_SEQ.DEFAUT_ACTIF    := FALSE;
GVL_SEQ.CODE_DEFAUT     := 0;

// ── Initialisation GVL_MOULES (stock initial terrain) ─────────
// CH1 AGADIR : N1=occupé(ID=1), N2=occupé(ID=1)
GVL_MOULES.CH[1,1].ID := 1;  GVL_MOULES.CH[1,1].OCCUPE := TRUE;
GVL_MOULES.CH[1,2].ID := 1;  GVL_MOULES.CH[1,2].OCCUPE := TRUE;
// CH2 IFRANE : N1=occupé(ID=2), N2=libre
GVL_MOULES.CH[2,1].ID := 2;  GVL_MOULES.CH[2,1].OCCUPE := TRUE;
GVL_MOULES.CH[2,2].ID := 0;  GVL_MOULES.CH[2,2].OCCUPE := FALSE;
// CH3 TANGER : N1=occupé(ID=3), N2=occupé(ID=3)
GVL_MOULES.CH[3,1].ID := 3;  GVL_MOULES.CH[3,1].OCCUPE := TRUE;
GVL_MOULES.CH[3,2].ID := 3;  GVL_MOULES.CH[3,2].OCCUPE := TRUE;
// CH4 RABAT : N1=occupé(ID=4), N2=occupé(ID=4)
GVL_MOULES.CH[4,1].ID := 4;  GVL_MOULES.CH[4,1].OCCUPE := TRUE;
GVL_MOULES.CH[4,2].ID := 4;  GVL_MOULES.CH[4,2].OCCUPE := TRUE;
// CH5 FEZ : N1=libre, N2=libre
GVL_MOULES.CH[5,1].ID := 0;  GVL_MOULES.CH[5,1].OCCUPE := FALSE;
GVL_MOULES.CH[5,2].ID := 0;  GVL_MOULES.CH[5,2].OCCUPE := FALSE;

GVL_MOULES.NB_EMPLACEMENTS_LIBRES := 3;
GVL_MOULES.MOULE_EN_PRESSE        := 0;

// ── Sécurité démarrage : toutes sorties physiques à FALSE ─────
GVL_IO.CMD_X_AV                := FALSE;
GVL_IO.CMD_X_AR                := FALSE;
GVL_IO.CMD_Z_HAUT              := FALSE;
GVL_IO.CMD_Z_BAS               := FALSE;
GVL_IO.CMD_SAT_EXT             := FALSE;
GVL_IO.CMD_SAT_RET             := FALSE;
GVL_IO.CMD_ROT_NORD            := FALSE;
GVL_IO.CMD_ROT_SUD             := FALSE;
GVL_IO.CMD_ARRET_PRESSE        := FALSE;
GVL_IO.CMD_DEBRIDAGE           := FALSE;
GVL_IO.CMD_BRIDAGE             := FALSE;
GVL_IO.CMD_AUTORISE_DEMARRAGE  := FALSE;
GVL_IO.CMD_MONTE_PILON         := FALSE;
GVL_IO.CMD_BAISSE_PILON        := FALSE;
GVL_IO.CMD_INTRO_ENTRE         := FALSE;
GVL_IO.CMD_INTRO_SORT          := FALSE;
GVL_IO.VOYANT_NETTOYAGE        := FALSE;
GVL_IO.BUZZER_DEBUT_NETTOYAGE  := FALSE;
GVL_IO.VOYANT_ATTENTE_ZONE_LIBRE := FALSE;

END_PROGRAM

(* ---- 18_PRG_MAIN.st ---- *)
// ================================================================
// 18_PRG_MAIN.st  —  Programme principal cyclique (équivalent OB1)
// CODESYS V3.5 — PROGRAM
// Configurer en tâche cyclique (ex : 10ms) dans le Task Manager
//
// Modification v2 — Laser OSSD :
//   - instLaser (FB_LaserSafe) ajouté : gère ZONE_CONFIRMEE automatiquement
//   - Ligne ZONE_CONFIRMEE manuelle supprimée (bouton remplacé par laser)
// ================================================================

PROGRAM PLC_PRG
VAR
    instG1    : FB_G1_Securite;
    instG0    : FB_G0_Conduite;
    instG2    : FB_G2_Homing;
    instG4    : FB_G4_AxeX;
    instG5    : FB_G5_AxeZ;
    instG6    : FB_G6_Rotation;
    instG7    : FB_G7_Satellite;
    instG8    : FB_G8_RFID;
    instG9    : FB_G9_Presse;
    instG10   : FB_G10_Intro;
    instG3    : FB_G3_Cycle;
    // ── IHM Visualization ────────────────────────────────────
    instHMI   : FB_HMI_Controller;
    instFault : FB_FaultInjector;
    // ── Sécurité laser OSSD (Sick S3000) ─────────────────────
    instLaser : FB_LaserSafe;
END_VAR

// ── IHM : textes, couleurs, boutons, injection défauts ────────
// Appel en premier : écrit dans GVL_IO avant les copies ci-dessous
instHMI();
instFault(
    FaultID   := GVL_HMI.HMI_FAULT_SEL,
    Inject    := GVL_HMI.HMI_BTN_INJECT,
    ResetFlt  := GVL_HMI.HMI_BTN_FAULT_RESET,
    Desc      => GVL_HMI.HMI_FAULT_DESC,
    Result    => GVL_HMI.HMI_FAULT_RESULT,
    FltActive => GVL_HMI.HMI_FAULT_ACTIVE
);

// ── Rafraîchissement commandes opérateur depuis GVL_IO ────────
GVL_SIG.OP_CMD_CM        := GVL_IO.CMD_CM;
GVL_SIG.OP_CMD_RESET     := GVL_IO.CMD_RESET;
GVL_SIG.OP_CMD_ACQ       := GVL_IO.CMD_ACQ_DEF;
GVL_SIG.OP_CMD_HOMING    := GVL_IO.CMD_HOMING_MANUEL;
GVL_SIG.OP_AU            := GVL_IO.AU_ACTIF;
GVL_SIG.OP_MOULE_DEMANDE := GVL_IO.MOULE_DEMANDE_HMI;
GVL_SIG.OP_MODE_AUTO     := GVL_IO.MODE_AUTO;
// ZONE_CONFIRMEE : géré par instLaser() ci-dessous — ne pas écrire ici
GVL_SIG.OP_PROLONG_NETTOYAGE := GVL_IO.PROLONG_NETTOYAGE_BTN OR GVL_HMI.HMI_BTN_PROLONG_NETTOYAGE;

// ── Images capteurs position X → GVL_SIG ─────────────────────
GVL_SIG.CAPTEUR_POS_X[0] := GVL_IO.POS_P0;
GVL_SIG.CAPTEUR_POS_X[1] := GVL_IO.POS_P1;
GVL_SIG.CAPTEUR_POS_X[2] := GVL_IO.POS_P2;
GVL_SIG.CAPTEUR_POS_X[3] := GVL_IO.POS_P3;
GVL_SIG.CAPTEUR_POS_X[4] := GVL_IO.POS_P4;
GVL_SIG.CAPTEUR_POS_X[5] := GVL_IO.POS_P5;
GVL_SIG.CAPTEUR_POS_X[6] := GVL_IO.POS_P6;

// ── Images présence chambres → GVL_SIG ───────────────────────
GVL_SIG.CAPTEUR_PRES_CH[1,1] := GVL_IO.CH1N1;
GVL_SIG.CAPTEUR_PRES_CH[1,2] := GVL_IO.CH1N2;
GVL_SIG.CAPTEUR_PRES_CH[2,1] := GVL_IO.CH2N1;
GVL_SIG.CAPTEUR_PRES_CH[2,2] := GVL_IO.CH2N2;
GVL_SIG.CAPTEUR_PRES_CH[3,1] := GVL_IO.CH3N1;
GVL_SIG.CAPTEUR_PRES_CH[3,2] := GVL_IO.CH3N2;
GVL_SIG.CAPTEUR_PRES_CH[4,1] := GVL_IO.CH4N1;
GVL_SIG.CAPTEUR_PRES_CH[4,2] := GVL_IO.CH4N2;
GVL_SIG.CAPTEUR_PRES_CH[5,1] := GVL_IO.CH5N1;
GVL_SIG.CAPTEUR_PRES_CH[5,2] := GVL_IO.CH5N2;

// ── Scanner laser OSSD — valide ZONE_CONFIRMEE automatiquement ─
// Doit être appelé AVANT instG3 pour que ZONE_CONFIRMEE soit à jour
instLaser();

// ── Appels GRAFCETs (ordre d'exécution fixe) ──────────────────
instG1();    // G1 Sécurité — EN PREMIER, toujours actif
instG0();    // G0 Superviseur modes
instG2();    // G2 Homing
instG4();    // G4 Axe X
instG5();    // G5 Axe Z
instG6();    // G6 Rotation
instG7();    // G7 Satellite
instG8();    // G8 RFID
instG9();    // G9 Presse
instG10();   // G10 Introducteur
instG3();    // G3 Cycle — EN DERNIER (coordinateur)

// ── Rafraîchissement voyants physiques depuis GVL_SIG ─────────
GVL_IO.VOYANT_MACHINE_PRETE  := GVL_SIG.VYT_MACHINE_PRETE;
GVL_IO.VOYANT_CYCLE_EN_COURS := GVL_SIG.VYT_CYCLE_EN_COURS;
GVL_IO.VOYANT_DEFAUT         := GVL_SIG.VYT_DEFAUT;
GVL_IO.VOYANT_INIT_OK        := GVL_SIG.VYT_INIT_OK;
GVL_IO.VOYANT_NETTOYAGE_TIMEOUT := GVL_SIG.VYT_NETTOYAGE_TIMEOUT;

END_PROGRAM

(* ---- 19_GVL_IO_HARDWARE_MAP.st ---- *)
// ================================================================
// 19_GVL_IO_HARDWARE_MAP.st
// CARTE COMPLÈTE I/O PHYSIQUES — ASRS QUADRA 10 / S7-1515
// Source : TIA_Import/Tags_ASRS.xml
//
// USAGE : Sur SoftPLC CODESYS (simulation) → utiliser GVL_IO sans AT
// USAGE : Sur automate physique → utiliser GVL avec AT %QX / %IX
//
// Pour activer les adresses hardware, remplacer dans GVL_IO.st :
//   CMD_X_AV : BOOL;
// par :
//   CMD_X_AV AT %QX0.0 : BOOL;
// ================================================================

// ── RÉSUMÉ ADRESSAGE SORTIES Q ────────────────────────────────
// %Q0.0   CMD_X_AV                Avance axe X
// %Q0.1   CMD_X_AR                Recul axe X
// %Q0.2   CMD_SAT_EXT             Extension satellite
// %Q0.3   CMD_SAT_RET             Rétraction satellite
// %Q0.4   CMD_Z_HAUT              Montée axe Z
// %Q0.5   CMD_Z_BAS               Descente axe Z
// %Q0.6   CMD_ROT_NORD            Rotation NORD
// %Q0.7   CMD_ROT_SUD             Rotation SUD
// %Q1.0   CMD_ARRET_PRESSE        Arrêt presse
// %Q1.1   CMD_DEBRIDAGE           Débridage moule
// %Q1.2   CMD_BRIDAGE             Bridage moule
// %Q1.3   CMD_AUTORISE_DEMARRAGE  Autorisation démarrage presse
// %Q1.4   CMD_MONTE_PILON         Montée pilon
// %Q1.5   CMD_BAISSE_PILON        Descente pilon
// %Q1.6   CMD_INTRO_ENTRE         Entrée introducteur ZPM
// %Q1.7   CMD_INTRO_SORT          Sortie introducteur ZPM
// %Q2.0   VOYANT_NETTOYAGE        Voyant nettoyage zone
// %Q2.1   BUZZER_DEBUT_NETTOYAGE  Buzzer début nettoyage
// %Q2.2   VOYANT_ATTENTE_ZONE_LIBRE
// %Q2.3   CMD_RFID_ACTIVER        Activation lecteur RFID RF350R
// %Q2.4   VOYANT_MACHINE_PRETE
// %Q2.5   VOYANT_CYCLE_EN_COURS
// %Q2.6   VOYANT_DEFAUT
// %Q2.7   VOYANT_INIT_OK
// %QW10   CONSIGNE_POS_X (WORD)   Consigne variateur axe X

// ── RÉSUMÉ ADRESSAGE ENTRÉES I ────────────────────────────────
// %I1.0   PRESSE_ARRETEE          Presse arrêtée confirmée
// %I1.1   MOULE_DEBRIDE           Moule débridé
// %I1.2   MOULE_BRIDE             Moule bridé
// %I1.3   PILON_HAUT_OK           Pilon en position haute
// %I1.4   PILON_BAS_OK            Pilon en position basse
// %I1.5   INTRODUCTEUR_EN_PRESSE  Introducteur en presse
// %I1.6   INTRODUCTEUR_A_ZPM      Introducteur à ZPM
// %I1.7   INTRO_VIDE              Introducteur vide
// %I2.0   MOULE_SUR_INTRO         Moule présent sur introducteur
// %I2.1   CAPTEUR_Z_TRANSPORT     Z position haute (transport)
// %I2.2   CAPTEUR_Z_NIVEAU1       Z niveau 1 chambre
// %I2.3   CAPTEUR_Z_NIVEAU2       Z niveau 2 chambre
// %I2.4   CAPTEUR_Z_ZPM           Z position ZPM
// %I2.5   CAPTEUR_CHARGE_CHARIOT  Charge présente sur fourches
// %I2.6   CAPTEUR_SAT_RETRACTE    Satellite rétracté
// %I2.7   CAPTEUR_SAT_ETENDU      Satellite étendu
// %I3.0   CAPTEUR_ZONE_OCCUPEE    Zone de travail occupée
// %I3.1   ZONE_LIBRE_BTN          Bouton zone libre opérateur
// %I3.2   CAPTEUR_ROT_NEUTRE      Rotation position neutre 0°
// %I3.3   CAPTEUR_ROT_NORD        Rotation position NORD
// %I3.4   CH1N1  Présence CH AGADIR N1
// %I3.5   CH1N2  Présence CH AGADIR N2
// %I3.6   CH2N1  Présence CH IFRANE N1
// %I3.7   CH2N2  Présence CH IFRANE N2
// %I4.0   CH3N1  Présence CH TANGER N1
// %I4.1   CH3N2  Présence CH TANGER N2
// %I4.2   CH4N1  Présence CH RABAT N1
// %I4.3   CH4N2  Présence CH RABAT N2
// %I4.4   CH5N1  Présence CH FEZ N1
// %I4.5   CH5N2  Présence CH FEZ N2
// %I4.6   RFID_LECTURE_OK         RFID lecture terminée
// %IB5    RFID_ID_LU (BYTE/USINT) ID moule lu par RFID MDS D160

// ── MERKERS M — COMMANDES HMI ─────────────────────────────────
// %M10.0  CMD_CM                  Commande changement moule
// %M10.1  CMD_RESET               Reset défaut
// %M10.2  CMD_ACQ_DEF             Acquittement défaut
// %M10.3  CMD_HOMING_MANUEL       Homing manuel
// %M10.4  AU_ACTIF                Arrêt urgence SW
// %M10.5  MODE_AUTO               Mode automatique
// %MB11   MOULE_DEMANDE_HMI       N° moule demandé (1-5)

// ── POSITIONS CAPTEURS X ──────────────────────────────────────
// (lire depuis Tags_ASRS.xml — adresses I5.x ou I6.x selon câblage)
// POS_P0..POS_P6 : capteurs de position chariot axe X

VAR_GLOBAL CONSTANT
    // Référence adresses pour documentation rapport
    ADDR_CMD_X_AV      : STRING := '%Q0.0';
    ADDR_CMD_Z_HAUT    : STRING := '%Q0.4';
    ADDR_PRESSE_ARRETEE: STRING := '%I1.0';
    ADDR_RFID_ID_LU    : STRING := '%IB5';
    ADDR_CMD_CM        : STRING := '%M10.0';
END_VAR
